// TIA Portal V21 export
// export: Created 2000-01-01T00:00:00.0000000Z, ExportSetting None
TYPE "UDT_HMI_FIO_Warehouse"
   STRUCT
      bExecuteCmd { ExternalWritable := 'False'} : Bool;   // HMI触发单次存取库作业（上升沿有效）
      bModeRetrieve { ExternalWritable := 'False'} : Bool;   // 作业模式：FALSE=入库(Store), TRUE=出库(Retrieve)
      bResetCmd { ExternalWritable := 'False'} : Bool;   // HMI故障复位命令
      iTargetCell { ExternalWritable := 'False'} : Int;   // HMI设定目标库位号 (1..54)
      tAxisSettleTime { ExternalWritable := 'False'} : Time;   // 升降/伸缩到位稳定延时（默认 T#800ms）
      tMoveTimeout { ExternalWritable := 'False'} : Time;   // 堆垛机寻址移动超时阈值（默认 T#10s）
      iCurrentStep { ExternalWritable := 'False'} : Int;   // 状态反馈：当前状态机步号
      iActiveTargetPos { ExternalWritable := 'False'} : Int;   // 状态反馈：当前输出给堆垛机的目标位置
      diStoredCount { ExternalWritable := 'False'} : DInt;   // 状态反馈：累计入库完成数
      diRetrievedCount { ExternalWritable := 'False'} : DInt;   // 状态反馈：累计出库完成数
      bBusy { ExternalWritable := 'False'} : Bool;   // 状态反馈：堆垛机作业忙
      bDone { ExternalWritable := 'False'} : Bool;   // 状态反馈：作业完成
      bFault { ExternalWritable := 'False'} : Bool;   // 状态反馈：故障标志
      wStatus { ExternalWritable := 'False'} : Word;   // 状态码：16#0000完成, 16#7000空闲, 16#7002执行中, 16#8200库位号越界, 16#8401动作超时, 16#8402急停触发
   END_STRUCT;
END_TYPE
